FUNCTION_BLOCK FB_Element_1 EXTENDS FB_SFC_Cycle IMPLEMENTS ITF_FB_SFC_Cycle
VAR_INPUT
	eElementID			: E_Element_List;

END_VAR
VAR_OUTPUT
END_VAR



VAR
	eType				: E_Element_Type;
	eProdType			: E_Product_Type;
	eState_Long			: E_Element_State_Long;
	eState_Short		: E_Element_State_Short;
	eState_Long_last	: E_Element_State_Long;
	eReq				: E_Request_List;
	eProcess			: E_Element_Process;




	i: INT;
	stStateChange		: TimeStruct;
	sState_Time			: STRING;
	
	sElementID			: STRING;
	eInterConnect		: E_InterConnection;
	bStataUpdate_Limited: BOOL;

	stCIP_Request: ST_CIP_Request;

	bTakePosInCIPBuffer_Partial: BOOL;
	bTakePosInCIPBuffer_Full: BOOL;
	bTakePosInCIPBuffer_Detergent: BOOL;
	bError: BOOL;
END_VAR

i:=i+1;
m_Set_SFCFlags_Reference();
SUPER^();
act_StateMachine();
act_StateChange_WatchGog();

sElementID:=TO_STRING(eElementID);

CASE eType OF 
	E_Element_Type.eTank:;
				act_Tank();
	E_Element_Type.eTriBlender:;
				act_TriBlender();
	E_Element_Type.eLine:;
				act_Line();

END_CASE

CASE eElementID OF
	E_Element_List.eTank_1:;
				eType:=E_Element_Type.eTank;
				eProdType:=E_Product_Type.Marinada;
				stCIP_Request.eClient:=E_CIP_Usage.eTank_1;
	E_Element_List.eTank_2:;
				eType:=E_Element_Type.eTank;
				eProdType:=E_Product_Type.Marinada;
				stCIP_Request.eClient:=E_CIP_Usage.eTank_2;
	E_Element_List.eTank_3:;
				eType:=E_Element_Type.eTank;
				eProdType:=E_Product_Type.Color;
				stCIP_Request.eClient:=E_CIP_Usage.eTank_3;
	E_Element_List.eTank_4:;
				eType:=E_Element_Type.eTank;
				eProdType:=E_Product_Type.Color;
				stCIP_Request.eClient:=E_CIP_Usage.eTank_4;
	E_Element_List.eTriBlender_Marinada:;
				eType:=E_Element_Type.eTriBlender;
				eProdType:=E_Product_Type.Marinada;		
				stCIP_Request.eClient:=E_CIP_Usage.eTriBlender_Marinada;
	E_Element_List.eTriBlender_Color:;
				eType:=E_Element_Type.eTriBlender;
				eProdType:=E_Product_Type.Color;
				stCIP_Request.eClient:=E_CIP_Usage.eTriBlender_Color;
	E_Element_List.eLine_Marinada:;
				eType:=E_Element_Type.eLine;
				eProdType:=E_Product_Type.Marinada;
				stCIP_Request.eClient:=E_CIP_Usage.eLine_Marinada;
	E_Element_List.eLine_Color:;
				eType:=E_Element_Type.eLine;
				eProdType:=E_Product_Type.Color;
				stCIP_Request.eClient:=E_CIP_Usage.eLine_Color;
END_CASE


IF bTakePosInCIPBuffer_Partial THEN;
	stCIP_Request.eType:=E_CIP_Type.R_Water;
	fbCIP.m_TakePosInCIPBuffer(stCIP_Request:=stCIP_Request);
	bTakePosInCIPBuffer_Partial:=FALSE;
END_IF

IF bTakePosInCIPBuffer_Detergent THEN;
	stCIP_Request.eType:=E_CIP_Type.Detergent;
	fbCIP.m_TakePosInCIPBuffer(stCIP_Request:=stCIP_Request);
	bTakePosInCIPBuffer_Detergent:=FALSE;
END_IF

IF bTakePosInCIPBuffer_Full THEN;
	stCIP_Request.eType:=E_CIP_Type.Full;
	fbCIP.m_TakePosInCIPBuffer(stCIP_Request:=stCIP_Request);
	bTakePosInCIPBuffer_Full:=FALSE;
END_IF

ACTION _aDone_entry:
eProcess:=E_Element_Process.eNone;
END_ACTION

ACTION _aInit_Tank_active:
SFCReset:=FALSE;
END_ACTION

ACTION _aInit_Tank_exit:
eProcess:=E_Element_Process.eNone;
END_ACTION

ACTION _aReady_active:


CASE eState_Long OF
	E_Element_State_Long.eOff,E_Element_State_Long.eStandby:;
			IF eReq=E_Request_List.eDrain THEN;
				eProcess:=E_Element_Process.eDrain;
			END_IF

	E_Element_State_Long.eCIP_5_Done:;
			IF eReq=E_Request_List.eWaterPrepare THEN;
				eProcess:=E_Element_Process.eFill_Water;
			END_IF	
			
	E_Element_State_Long.eWaterReady:;
			IF eReq=E_Request_List.eDissolve THEN;
				eProcess:=E_Element_Process.eDissolving;
			END_IF	

	E_Element_State_Long.eReady:;
			IF eReq=E_Request_List.eProduction THEN;
				eProcess:=E_Element_Process.eConnectionToLine;
			END_IF	

	E_Element_State_Long.eProduction:;
			IF eReq=E_Request_List.eDisconnectTank THEN;
				eProcess:=E_Element_Process.eDisconnection;
			END_IF			

END_CASE
END_ACTION

ACTION _aState_Update_01_entry:
eState_Long:=E_Element_State_Long.eNotClean;
END_ACTION

ACTION _aState_Update_02_entry:
eState_Long:=E_Element_State_Long.eWaterReady;
END_ACTION

ACTION _aState_Update_03_entry:
eState_Long:=E_Element_State_Long.eReady;
END_ACTION

ACTION _aState_Update_04_entry:
eState_Long:=E_Element_State_Long.eProduction;
END_ACTION

ACTION _aState_Update_05_entry:
eState_Long:=E_Element_State_Long.eReady;
END_ACTION

ACTION act_Line:

END_ACTION

ACTION act_Oper_Tank:
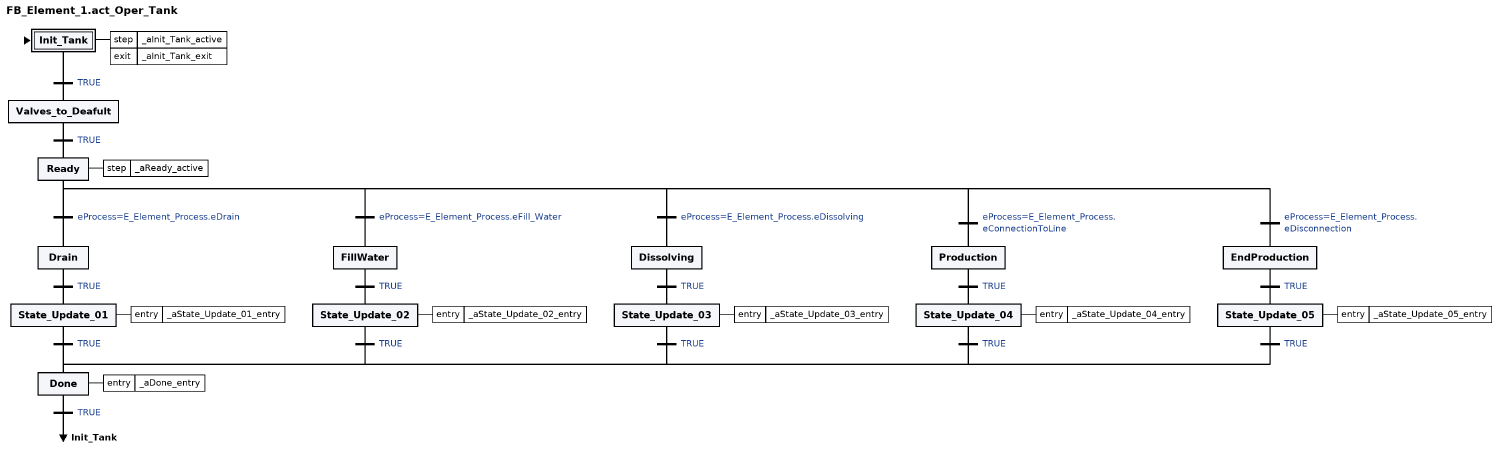
INITIAL_STEP Init_Tank:  // min time T#2s
    _aInit_Tank_active(N);  // step action
    _aInit_Tank_exit(P0);  // exit action
END_STEP
TRANSITION FROM Init_Tank TO Valves_to_Deafult
    := TRUE;
END_TRANSITION
STEP Valves_to_Deafult:
END_STEP
TRANSITION FROM Valves_to_Deafult TO Ready
    := TRUE;
END_TRANSITION
STEP Ready:  // min time T#2s
    _aReady_active(N);  // step action
END_STEP
TRANSITION FROM Ready TO Drain
    := eProcess=E_Element_Process.eDrain;
END_TRANSITION
STEP Drain:
END_STEP
TRANSITION FROM Drain TO State_Update_01
    := TRUE;
END_TRANSITION
STEP State_Update_01:
    _aState_Update_01_entry(P1);  // entry action
END_STEP
TRANSITION FROM State_Update_01 TO Done
    := TRUE;
END_TRANSITION
TRANSITION FROM Ready TO FillWater
    := eProcess=E_Element_Process.eFill_Water;
END_TRANSITION
STEP FillWater:
END_STEP
TRANSITION FROM FillWater TO State_Update_02
    := TRUE;
END_TRANSITION
STEP State_Update_02:
    _aState_Update_02_entry(P1);  // entry action
END_STEP
TRANSITION FROM State_Update_02 TO Done
    := TRUE;
END_TRANSITION
TRANSITION FROM Ready TO Dissolving
    := eProcess=E_Element_Process.eDissolving;
END_TRANSITION
STEP Dissolving:
END_STEP
TRANSITION FROM Dissolving TO State_Update_03
    := TRUE;
END_TRANSITION
STEP State_Update_03:
    _aState_Update_03_entry(P1);  // entry action
END_STEP
TRANSITION FROM State_Update_03 TO Done
    := TRUE;
END_TRANSITION
TRANSITION FROM Ready TO Production
    := eProcess=E_Element_Process.eConnectionToLine;
END_TRANSITION
STEP Production:
END_STEP
TRANSITION FROM Production TO State_Update_04
    := TRUE;
END_TRANSITION
STEP State_Update_04:
    _aState_Update_04_entry(P1);  // entry action
END_STEP
TRANSITION FROM State_Update_04 TO Done
    := TRUE;
END_TRANSITION
TRANSITION FROM Ready TO EndProduction
    := eProcess=E_Element_Process.eDisconnection;
END_TRANSITION
STEP EndProduction:
END_STEP
TRANSITION FROM EndProduction TO State_Update_05
    := TRUE;
END_TRANSITION
STEP State_Update_05:
    _aState_Update_05_entry(P1);  // entry action
END_STEP
TRANSITION FROM State_Update_05 TO Done
    := TRUE;
END_TRANSITION
STEP Done:  // min time T#2s
    _aDone_entry(P1);  // entry action
END_STEP
TRANSITION FROM Done TO Init_Tank
    := TRUE;
END_TRANSITION
// branch label Branch0_act_Oper_Tank
END_ACTION

ACTION act_StateChange_WatchGog:
IF eState_Long<>eState_Long_last THEN;
	eState_Long_last:=eState_Long;
	stStateChange:=stSystemTime;
END_IF

sState_Time:=prg_RealClock.m_DeltaTime(stStartTime:=stStateChange);
END_ACTION

ACTION act_StateMachine:


CASE eState_Long OF
	E_Element_State_Long.eOff,
	E_Element_State_Long.eStandby,
	E_Element_State_Long.eNotClean,
	E_Element_State_Long.eCIP_1_Rinzed,
	E_Element_State_Long.eCIP_2_Deterged,
	E_Element_State_Long.eCIP_3_Deterged_Clean,	
	E_Element_State_Long.eCIP_4_Sanitized:;
				eState_Short:=E_Element_State_Short.eNotClean;

	E_Element_State_Long.eCIP_5_Done,	
	E_Element_State_Long.eWaterReady:;	
				eState_Short:=E_Element_State_Short.eClean;

	E_Element_State_Long.eReady,
	E_Element_State_Long.eProduction,
	E_Element_State_Long.eEmpty,	
	E_Element_State_Long.eExpired:;
				eState_Short:=E_Element_State_Short.eProduct;
	
END_CASE
END_ACTION

ACTION act_Tank:
act_Oper_Tank();
END_ACTION

ACTION act_TriBlender:
IF eInterConnect=E_InterConnection.ConnToCIP 
AND eElementID=E_Element_List.eTriBlender_Marinada
AND eTriBlenderPipe<>E_TriBlenderPipe.eMarinada
THEN;
	bError:=TRUE;
ELSE;
	bError:=FALSE;
END_IF
END_ACTION

METHOD m_Disconnect : BOOL
VAR_INPUT
END_VAR
eInterConnect:=E_InterConnection.NotConnected;
//bInterConnectedToLine:=FALSE;
END_METHOD

METHOD m_InterConnect : BOOL
VAR_INPUT
	value: E_InterConnection;
END_VAR
eInterConnect:=value;
END_METHOD

METHOD m_InterConnected_State : BOOL
VAR_INPUT
	eState_Long_Set			: E_Element_State_Long;
END_VAR

IF eState_Long_Set>eState_Long 
OR eState_Long_Set=E_Element_State_Long.eNotClean
THEN;
	eState_Long:=eState_Long_Set;
END_IF
END_METHOD

METHOD m_Set_SFCFlags_Reference : BOOL
//Set reference to SFC flags

refSFC.SFCInit REF= SFCInit;
refSFC.SFCReset REF= SFCReset;
refSFC.SFCError REF= SFCError;
refSFC.SFCEnableLimit REF= SFCEnableLimit;
refSFC.SFCErrorStep REF= SFCErrorStep;
refSFC.SFCErrorPOU REF= SFCErrorPOU;
refSFC.SFCQuitError REF= SFCQuitError;
refSFC.SFCPause REF= SFCPause;
refSFC.SFCTrans REF= SFCTrans;
refSFC.SFCCurrentStep REF= SFCCurrentStep;
refSFC.SFCTip REF= SFCTip;
refSFC.SFCTipMode REF= SFCTipMode;

// Cycle handle for SFC
m_SFC_Handle();
END_METHOD

METHOD m_StateUpdate_Limit : BOOL
VAR_INPUT
	value: BOOL;
END_VAR
IF value THEN;
	bStataUpdate_Limited:=TRUE;
ELSE;
	bStataUpdate_Limited:=FALSE;
END_IF
END_METHOD

END_FUNCTION_BLOCK

(* stored: Version 1.1.0.1, ProductVersion 3.1.4024.12
   POU FB_Element_1: Id {0c9cbe8c-7dda-4561-8ed0-d554091062a9}, SpecialFunc None
   Folder Manage: Id {f254e61f-7e1a-4990-bdd7-86e543689a33}
   Action _aDone_entry: Id {f360ca42-d94b-4deb-84bc-6f864703f808}
   Action _aInit_Tank_active: Id {c45b88da-7ee2-4ff7-b069-9b4e0aa4c520}
   Action _aInit_Tank_exit: Id {0d4569d4-ff75-48f1-9c70-281e68ef9a3f}
   Action _aReady_active: Id {06b27a2a-0dd3-4a72-b37c-f884be26cb36}
   Action _aState_Update_01_entry: Id {1b8601ca-09e9-4f2c-82b5-44f30e8ef1a2}
   Action _aState_Update_02_entry: Id {b77f594f-e63c-47e5-953b-38b9889ddafb}
   Action _aState_Update_03_entry: Id {82ddc7d9-7cfa-4429-80f4-755528c1e2ef}
   Action _aState_Update_04_entry: Id {53585974-6ceb-4a8b-abcd-a407e5f278a9}
   Action _aState_Update_05_entry: Id {7631ace1-468f-40fd-8d9e-d215e3c98e12}
   Action act_Line: Id {0ec62730-e61a-41a2-924c-51671604578b}
   Action act_Oper_Tank: Id {7dde56e5-1f54-43e6-9270-d42adcb20fc5}
   Action act_StateChange_WatchGog: Id {c16d49dc-334d-49fe-813a-17142978f429}
   Action act_StateMachine: Id {b706c936-cbcf-4a3a-9be1-20180bdd8aa1}
   Action act_Tank: Id {6200ac69-7f3b-413b-a098-3397c80ffe69}
   Action act_TriBlender: Id {16b91cbd-73ec-4a6a-930a-0161124493e4}
   Method m_Disconnect: Id {f6370718-b114-4e04-a5b7-17ebbef5b212}
   Method m_InterConnect: Id {297c1053-5f16-4296-99d3-3cca348c0902}
   Method m_InterConnected_State: Id {47b4c791-7b17-48f2-9da1-481769db6a71}
   Method m_Set_SFCFlags_Reference: Id {843fc4cc-8e41-43dd-8aa7-4e962c29228c}
   Method m_StateUpdate_Limit: Id {100144a5-3c55-4e4c-8c08-914b0d81d778} *)
